(* IEC 61131-3 sources: Lasal-MCP/examples/SampleSource/LASALScreenAdvancedSolution/LASALScreenAdvancedSolution/LASALScreenAdvacnedSolution/Stations/Terminal/HMI/Class/DataRecordFileHandling, 1 file *)

(* ---- DataRecordFileHandling.st ---- *)
(*!
<Class
	Name               = "DataRecordFileHandling"
	Revision           = "0.0"
	RealtimeTask       = "false"
	CyclicTask         = "false"
	BackgroundTask     = "true"
	DefBackground      = "50 ms"
	Sigmatek           = "false"
	OSInterface        = "false"
	HighPriority       = "false"
	Automatic          = "false"
	UpdateMode         = "Prescan"
	SharedCommandTable = "true"
	Objectsize         = "(720,180)">
	<Channels>
		<Server Name="DriveName" Visualized="true" Remotely="true" Initialize="true" WriteProtected="false" Retentive="false"/>
		<Server Name="FileExtension" Visualized="true" Remotely="true" Initialize="true" WriteProtected="false" Retentive="false"/>
		<Server Name="FileIsCreated" Visualized="false" Initialize="false" WriteProtected="true" Retentive="false"/>
		<Server Name="FileName" Visualized="true" Remotely="true" Initialize="true" WriteProtected="false" Retentive="false"/>
		<Server Name="IntError" Visualized="false" Initialize="false" WriteProtected="true" Retentive="false"/>
		<Server Name="StartFileWrite" Visualized="false" Initialize="false" WriteProtected="false" Retentive="false"/>
		<Server Name="Steps" Visualized="false" Initialize="false" WriteProtected="true" Retentive="false"/>
		<Client Name="_FileSys" Required="false" Internal="false"/>
		<Client Name="DataRecordFileRead" Required="true" Internal="false"/>
		<Client Name="DriveNameString" Required="true" Internal="true"/>
		<Client Name="FileExtensionString" Required="true" Internal="true"/>
		<Client Name="FileNameString" Required="true" Internal="true"/>
		<Client Name="SigCLib" Required="false" Internal="false"/>
	</Channels>
	<Network Name="DataRecordFileHandling">
		<!-- List of Components in this network -->
		<Components>
			<Object
				Name       = "DriveNameString"
				Class      = "StringRAM"
				Position   = "(60,390)"
				Visualized = "true"
				Remotely   = "true">
				<Channels>
					<Server Name="Data"/>
					<Client Name="SingleRealloc" Value="1"/>
					<Client Name="UseFile"/>
				</Channels>
			</Object>
			<Object
				Name       = "FileExtensionString"
				Class      = "StringRAM"
				Position   = "(60,810)"
				Visualized = "true"
				Remotely   = "true">
				<Channels>
					<Server Name="Data"/>
					<Client Name="SingleRealloc" Value="1"/>
					<Client Name="UseFile"/>
				</Channels>
			</Object>
			<Object
				Name       = "FileNameString"
				Class      = "StringRAM"
				Position   = "(60,600)"
				Visualized = "true"
				Remotely   = "true">
				<Channels>
					<Server Name="Data"/>
					<Client Name="SingleRealloc" Value="1"/>
					<Client Name="UseFile"/>
				</Channels>
			</Object>
		</Components>
		<Comments>
		</Comments>
		<!-- List of Connections in this network -->
		<Connections>
			<Connection Source="this.DriveNameString" Destination="DriveNameString.Data"/>
			<Connection Source="this.FileNameString" Destination="FileNameString.Data"/>
			<Connection Source="this.FileExtensionString" Destination="FileExtensionString.Data"/>
			<Connection Source="this.DriveName" Destination="DriveNameString.Data" Vertices="(728,450),(556,480),"/>
			<Connection Source="this.FileName" Destination="FileNameString.Data" Vertices="(728,510),(556,690),"/>
			<Connection Source="this.FileExtension" Destination="FileExtensionString.Data" Vertices="(728,570),(556,900),"/>
		</Connections>
		<!-- Headerfiles -->
		<Options>
		</Options>
	</Network>
</Class>
*)
DataRecordFileHandling : CLASS
	TYPE
	  _FILE_STEPS :  //! <Type Public="true" Name="_FILE_STEPS"/>
	  (
	    FS_Idle,
	    FS_FileCreate,
	    FS_WaitFileCreated,
	    FS_FileClose,
	    FS_WaitFileClosed,
	    FS_FileOpen,
	    FS_WaitFileOpened,
	    FS_FileWrite,
	    FS_WaitFileWritten,
	    FS_FileLength,
	    FS_WaitFileLength,
	    FS_Error
	  )$UDINT;
	END_TYPE
  //Servers:
	Steps 	: SvrChCmd__FILE_STEPS_PTofCls_DataRecordFileHandling;
	StartFileWrite 	: SvrCh_DINT;
	FileIsCreated 	: SvrCh_DINT;
	IntError 	: SvrCh_DINT;
	DriveName 	: SvrCh_UDINT;
	FileName 	: SvrCh_UDINT;
	FileExtension 	: SvrCh_UDINT;
  //Clients:
	_FileSys 	: CltChCmd__FileSys;
	SigCLib 	: CltChCmd_SigCLib;
	DataRecordFileRead 	: CltChCmd_DataRecordFileRead;
	DriveNameString 	: CltChCmd_StringRAM;
	FileNameString 	: CltChCmd_StringRAM;
	FileExtensionString 	: CltChCmd_StringRAM;
  //Variables:
		TempFullFileName : ARRAY [0..255] OF CHAR;

		FileHandle 	: DINT;
		AsyncId 	: DINT;
		Length 	: UDINT;
		pSaveData 	: ^DINT;
		FileIsRead 	: BOOL;
  //Functions:

	FUNCTION VIRTUAL GLOBAL Init;

	FUNCTION VIRTUAL GLOBAL Background
		VAR_INPUT
			EAX 	: UDINT;
		END_VAR
		VAR_OUTPUT
			state (EAX) 	: UDINT;
		END_VAR;

	FUNCTION GLOBAL StartWrite
		VAR_INPUT
			pData 	: ^DINT;
			Amount 	: UDINT;
		END_VAR
		VAR_OUTPUT
			Retcode 	: DINT;
		END_VAR;

	FUNCTION VIRTUAL GLOBAL DriveName::Read
		VAR_OUTPUT
			output (EAX) 	: UDINT;
		END_VAR;

	FUNCTION VIRTUAL GLOBAL DriveName::Write
		VAR_INPUT
			input (EAX) 	: UDINT;
		END_VAR
		VAR_OUTPUT
			result (EAX) 	: UDINT;
		END_VAR;

	FUNCTION VIRTUAL GLOBAL FileName::Read
		VAR_OUTPUT
			output (EAX) 	: UDINT;
		END_VAR;

	FUNCTION VIRTUAL GLOBAL FileName::Write
		VAR_INPUT
			input (EAX) 	: UDINT;
		END_VAR
		VAR_OUTPUT
			result (EAX) 	: UDINT;
		END_VAR;

	FUNCTION VIRTUAL GLOBAL FileExtension::Read
		VAR_OUTPUT
			output (EAX) 	: UDINT;
		END_VAR;

	FUNCTION VIRTUAL GLOBAL FileExtension::Write
		VAR_INPUT
			input (EAX) 	: UDINT;
		END_VAR
		VAR_OUTPUT
			result (EAX) 	: UDINT;
		END_VAR;
  //Tables:
	FUNCTION @STD
		VAR_OUTPUT
			ret_code	: CONFSTATES;
		END_VAR;
	FUNCTION GLOBAL TAB @CT_;
END_CLASS;

#pragma using StringRAM
#pragma usingLtd _FileSys
#pragma usingLtd DataRecordFileRead
#pragma usingLtd SigCLib

FUNCTION VIRTUAL GLOBAL DataRecordFileHandling::Init

  if (_FirstScan = TRUE) then
    Steps := FS_FileCreate; // Create file in the beginning
  end_if;

END_FUNCTION

FUNCTION VIRTUAL GLOBAL DataRecordFileHandling::Background
	VAR_INPUT
		EAX 	: UDINT;
	END_VAR
	VAR_OUTPUT
		state (EAX) 	: UDINT;
	END_VAR
  VAR
    locBuffer : ARRAY[0..255] of CHAR;
    stringLength : UDINT;
    pError : ^CHAR;
    fileWritten : DINT;
    asyncState : DINT;
  END_VAR

  // ==========================================================================
  case Steps of
    // --------------------------------------------------------------
  	FS_Idle:

      if (StartFileWrite = 1) then
        StartFileWrite := 0;
        Steps := FS_FileOpen;
      end_if;

    // --------------------------------------------------------------
  	FS_FileCreate:

      // Get drive name
      stringLength := DriveNameString.GetLength();

      DriveNameString.GetDataAt(pData:= #locBuffer[0],
                                udSize:= stringLength,
                                udAt:= 0);

      locBuffer[stringLength] := 0;

      pError := SigCLib.StrCpy(dst0:= #TempFullFileName[0],
                               src0:= #locBuffer[0]);

      if (pError <> #TempFullFileName[0]) then
        IntError := -1;
        Steps := FS_Error;
        return;
      end_if;

      // Get file name
      stringLength := FileNameString.GetLength();

      FileNameString.GetDataAt(pData:= #locBuffer[0],
                         udSize:= stringLength,
                         udAt:= 0);

      locBuffer[stringLength] := 0;

      pError := SigCLib.StrCat(ps1:= #TempFullFileName[0],
                               ps2:= #locBuffer[0]);

      if (pError <> #TempFullFileName[0]) then
        IntError := -2;
        Steps := FS_Error;
        return;
      end_if;

      // Get file extension
      stringLength := FileExtensionString.GetLength();

      FileExtensionString.GetDataAt(pData:= #locBuffer[0],
                                    udSize:= stringLength,
                                    udAt:= 0);

      locBuffer[stringLength] := 0;

      pError := SigCLib.StrCat(ps1:= #TempFullFileName[0],
                               ps2:= #locBuffer[0]);

      if (pError <> #TempFullFileName[0]) then
        IntError := -3;
        Steps := FS_Error;
        return;
      end_if;

      AsyncId := _FileSys.FileCreate_A(Async:= 1,
                                       dpne:= #TempFullFileName[0],
                                       size:= 1 MB,
                                       fill:= 0,
                                       att:= ATT_CREATE_ALWAYS);

      Steps := FS_WaitFileCreated;

    // --------------------------------------------------------------
  	FS_WaitFileCreated:

      asyncState := _FileSys.GetAsyncState(ID:= to_udint(AsyncId),
                                           Erg:= #FileHandle);

      // ==================================================
      case asyncState of
        //---------------------------------------
        0:
          if (FileHandle >= 0) then
            Steps := FS_FileClose;
          else
            IntError := -4;
            Steps := FS_Error;
          end_if;

        //---------------------------------------
        RT_ERG_DELETED,
        RT_INVALID_ID:
          IntError := -5;
          Steps := FS_Error;

        //---------------------------------------
        RT_NOT_STARTED,
        RT_IN_PROGRESS:

      end_case;
      // ==================================================

    // --------------------------------------------------------------
  	FS_FileClose:

      AsyncId := _FileSys.FileClose_A(Async:= 1,
                                      handle:= FileHandle);

      Steps := FS_WaitFileClosed;

    // --------------------------------------------------------------
  	FS_WaitFileClosed:

      asyncState := _FileSys.GetAsyncState(ID:= to_udint(AsyncId),
                                           Erg:= #FileHandle);

      // ==================================================
      case asyncState of
        //---------------------------------------
        0:
          if (FileHandle >= 0) then
            if FileIsCreated then
              Steps := FS_Idle;
            else
              FileIsCreated := 1;
              Steps := FS_FileOpen;
            end_if;
          else
            IntError := -6;
            Steps := FS_Error;
          end_if;

        //---------------------------------------
        RT_ERG_DELETED,
        RT_INVALID_ID:
          IntError := -7;
          Steps := FS_Error;

        //---------------------------------------
        RT_NOT_STARTED,
        RT_IN_PROGRESS:

      end_case;
      // ==================================================

    // --------------------------------------------------------------
  	FS_FileOpen:

      AsyncId := _FileSys.FileOpen_A(Async:= 1,
                                     FileName:= #TempFullFileName[0],
                                     attributes:= ATT_READ_WRITE);

      Steps := FS_WaitFileOpened;

    // --------------------------------------------------------------
  	FS_WaitFileOpened:

      asyncState := _FileSys.GetAsyncState(ID:= to_udint(AsyncId),
                                           Erg:= #FileHandle);

      // ==================================================
      case asyncState of
        //---------------------------------------
        0:
          if (FileHandle >= 0) then

            Steps := FS_FileWrite;

          elsif FileHandle = -16 then
            Steps := FS_FileCreate;
          else
            IntError := -8;
            Steps := FS_Error;
          end_if;

        //---------------------------------------
        RT_ERG_DELETED,
        RT_INVALID_ID:
          IntError := -9;
          Steps := FS_Error;

        //---------------------------------------
        RT_NOT_STARTED,
        RT_IN_PROGRESS:

      end_case;
      // ==================================================

    // --------------------------------------------------------------
  	FS_FileWrite:

      AsyncId := _FileSys.FileWrite_A(Async:= 1,
                                      handle:= FileHandle,
                                      buffer:= pSaveData,
                                      Length:= Length);

      Steps := FS_WaitFileWritten;

    // --------------------------------------------------------------
  	FS_WaitFileWritten:

      asyncState := _FileSys.GetAsyncState(ID:= to_udint(AsyncId),
                                           Erg:= #fileWritten);

      // ==================================================
      case asyncState of
        //---------------------------------------
        0:
          if (fileWritten >= 0) then
            Steps := FS_FileClose;
          else
            IntError := -10;
            Steps := FS_Error;
          end_if;

        //---------------------------------------
        RT_ERG_DELETED,
        RT_INVALID_ID:
          IntError := -11;
          Steps := FS_Error;

        //-----------------------------------
        RT_NOT_STARTED,
        RT_IN_PROGRESS:

      end_case;
      // ==================================================

    // --------------------------------------------------------------
    FS_Error:

  end_case;
  // ==========================================================================

	state := READY;

END_FUNCTION

FUNCTION VIRTUAL GLOBAL DataRecordFileHandling::DriveName::Read
	VAR_OUTPUT
		output (EAX) 	: UDINT;
	END_VAR

	DriveName := DriveNameString.Data.Read();
	output := DriveName;

END_FUNCTION

FUNCTION VIRTUAL GLOBAL DataRecordFileHandling::DriveName::Write
	VAR_INPUT
		input (EAX) 	: UDINT;
	END_VAR
	VAR_OUTPUT
		result (EAX) 	: UDINT;
	END_VAR

	DriveName := input;
	result := (DriveNameString.Data.Write(DriveName))$UDINT;

END_FUNCTION

FUNCTION VIRTUAL GLOBAL DataRecordFileHandling::FileName::Read
	VAR_OUTPUT
		output (EAX) 	: UDINT;
	END_VAR

	FileName := FileNameString.Data.Read();
	output := FileName;

END_FUNCTION

FUNCTION VIRTUAL GLOBAL DataRecordFileHandling::FileName::Write
	VAR_INPUT
		input (EAX) 	: UDINT;
	END_VAR
	VAR_OUTPUT
		result (EAX) 	: UDINT;
	END_VAR

	FileName := input;
	result := (FileNameString.Data.Write(FileName))$UDINT;

END_FUNCTION

FUNCTION VIRTUAL GLOBAL DataRecordFileHandling::FileExtension::Read
	VAR_OUTPUT
		output (EAX) 	: UDINT;
	END_VAR

	FileExtension := FileExtensionString.Data.Read();
	output := FileExtension;

END_FUNCTION

FUNCTION VIRTUAL GLOBAL DataRecordFileHandling::FileExtension::Write
	VAR_INPUT
		input (EAX) 	: UDINT;
	END_VAR
	VAR_OUTPUT
		result (EAX) 	: UDINT;
	END_VAR

	FileExtension := input;
	result := (FileExtensionString.Data.Write(FileExtension))$UDINT;

END_FUNCTION

FUNCTION GLOBAL DataRecordFileHandling::StartWrite
	VAR_INPUT
		pData 	: ^DINT;
		Amount 	: UDINT;
	END_VAR
	VAR_OUTPUT
		Retcode 	: DINT;
	END_VAR

  if (pData = NIL) then
    IntError := -14;
    Retcode := -1;
    return;
  end_if;

  if (FileIsCreated = 0) then
    Retcode := -2;
    return;
  end_if;

  pSaveData := pData;
  Length := Amount;
  FileIsRead := FALSE;
  Steps := FS_FileOpen;

END_FUNCTION
